Staubli VAL3: BP_Validation.pgx

program BP_Validation()
begin
  bStart[0] = true
end
